Fanuc KAREL source: KT00981.KL

PROGRAM KT00981
%NOLOCKGROUP
VAR
  I1: INTEGER
  I2: INTEGER
  CFG: CONFIG
  OUT: XYZWPREXT
BEGIN
  I1 = 2
  I2 = 3
  I1 = 2
  I2 = 3
  CFG.CFG_FLIP = TRUE
  OUT = POS(I1, I1, I1, I1, I1, I1, CFG)
END KT00981
